Fanuc KAREL source: KO00110.KL

PROGRAM KO00110
%NOLOCKGROUP
VAR
  A: REAL
  B: ARRAY[2] OF BYTE
  OUT: REAL
BEGIN
  A = 1
  B[1] = 2
  OUT = ATAN2(A, B[1])
END KO00110
